(*
SPDX-FileCopyrightText: © 2026 Oleksandr Tiutyk <trofimich@gmail.com>
SPDX-License-Identifier: MIT
License: https://opensource.org/license/mit
*)

(*!
<summary>Provides static helper methods for throwing Workflow-specific exceptions.</summary>
<description>
Constructs stack-local template exceptions, formats diagnostics without heap allocation and propagates them
through ExceptionManager. Formatting uses bounded storage; propagation may allocate a registered clone.
Call only from cyclic execution, outside lifecycle methods. Each template is call-local; exception ownership
and task-boundary cleanup remain governed by Core.ExceptionManager and DynamicMemoryManager.
</description>
*)

{attribute 'no_explicit_call' := 'do not call this function block directly'}
PROGRAM WorkflowExceptions
VAR
	{attribute 'hide'} 
	_ClassName : STRING := __POUNAME();
END_VAR

(*!
<summary>Returns the diagnostic name stored by this program.</summary>
<description>
Borrows program-owned storage. Treat the returned reference as read-only and do not use it to change metadata.
</description>
*)
{attribute 'monitoring' := 'call'}
PROPERTY ClassName : REFERENCE TO STRING
GET
ClassName REF= _ClassName;
END_GET
END_PROPERTY

(*!
<summary>Returns the compiler-initialized library namespace.</summary>
<description>
Borrows shared read-only namespace storage; no allocation or ownership transfer occurs.
</description>
*)
{attribute 'monitoring' := 'call'}
PROPERTY NamespaceName : REFERENCE TO STRING
GET
NamespaceName REF= CurrentNamespace.Name;
END_GET
END_PROPERTY

(*!
<summary>Raises an InvalidNestedWorkflowStateException without requiring a caller-owned exception variable.</summary>
<description>
Constructs a temporary stack template and delegates to InvalidNestedWorkflowStateException.Throw.
</description>
<param name="sourceNamespaceName">Namespace of the caller.</param>
<param name="sourceClassName">Class name of the caller.</param>
<param name="sourcePOUName">POU name of the caller.</param>
<param name="sourcePosition">Source position of the caller.</param>
<param name="nestedActivityState">Observed child workflow element state.</param>
*)
METHOD ThrowInvalidNestedWorkflowState
VAR_INPUT
	sourceNamespaceName : STRING;
	sourceClassName : STRING;
	sourcePOUName : STRING;
	sourcePosition : STRING;
	nestedActivityState : WORKFLOW_ELEMENT_STATE;
END_VAR
VAR
	exception : InvalidNestedWorkflowStateException;
END_VAR
exception.Throw(
	sourceNamespaceName := sourceNamespaceName,
	sourceClassName := sourceClassName,
	sourcePOUName := sourcePOUName,
	sourcePosition := sourcePosition,
	nestedActivityState := nestedActivityState
);
END_METHOD

(*!
<summary>Raises an InvalidWorkflowTransitionException without requiring a caller-owned exception variable.</summary>
<description>
Constructs a temporary stack template and delegates to InvalidWorkflowTransitionException.Throw.
</description>
<param name="sourceNamespaceName">Namespace of the caller.</param>
<param name="sourceClassName">Class name of the caller.</param>
<param name="sourcePOUName">POU name of the caller.</param>
<param name="sourcePosition">Source position of the caller.</param>
<param name="fromState">Current state of the workflow element.</param>
<param name="toState">Rejected target state.</param>
*)
METHOD ThrowInvalidWorkflowTransition
VAR_INPUT
	sourceNamespaceName : STRING;
	sourceClassName : STRING;
	sourcePOUName : STRING;
	sourcePosition : STRING;
	fromState : WORKFLOW_ELEMENT_STATE;
	toState : WORKFLOW_ELEMENT_STATE;
END_VAR
VAR
	exception : InvalidWorkflowTransitionException;
END_VAR
exception.Throw(
	sourceNamespaceName := sourceNamespaceName,
	sourceClassName := sourceClassName,
	sourcePOUName := sourcePOUName,
	sourcePosition := sourcePosition,
	fromState := fromState,
	toState := toState
);
END_METHOD

(*!
<summary>Raises a WorkflowAttachmentException without requiring a caller-owned exception variable.</summary>
<description>Constructs a temporary stack template and delegates to WorkflowAttachmentException.Throw.</description>
<param name="sourceNamespaceName">Namespace of the caller.</param>
<param name="sourceClassName">Class name of the caller.</param>
<param name="sourcePOUName">POU name of the caller.</param>
<param name="sourcePosition">Source position of the caller.</param>
<param name="message">Diagnostic explanation.</param>
*)
METHOD ThrowWorkflowAttachment
VAR_INPUT
	sourceNamespaceName : STRING;
	sourceClassName : STRING;
	sourcePOUName : STRING;
	sourcePosition : STRING;
END_VAR
VAR_IN_OUT CONSTANT
	message : TOF_Core.ERROR_MESSAGE;
END_VAR
VAR
	exception : WorkflowAttachmentException;
END_VAR
exception.Throw(
	sourceNamespaceName := sourceNamespaceName,
	sourceClassName := sourceClassName,
	sourcePOUName := sourcePOUName,
	sourcePosition := sourcePosition,
	message := message
);
END_METHOD

(*!
<summary>Raises a WorkflowConfigurationException without requiring a caller-owned exception variable.</summary>
<description>Constructs a temporary stack template and delegates to WorkflowConfigurationException.Throw.</description>
<param name="sourceNamespaceName">Namespace of the caller.</param>
<param name="sourceClassName">Class name of the caller.</param>
<param name="sourcePOUName">POU name of the caller.</param>
<param name="sourcePosition">Source position of the caller.</param>
<param name="message">Diagnostic explanation.</param>
*)
METHOD ThrowWorkflowConfiguration
VAR_INPUT
	sourceNamespaceName : STRING;
	sourceClassName : STRING;
	sourcePOUName : STRING;
	sourcePosition : STRING;
	message : WSTRING(255);
END_VAR
VAR
	exception : WorkflowConfigurationException;
END_VAR
exception.Throw(
	sourceNamespaceName := sourceNamespaceName,
	sourceClassName := sourceClassName,
	sourcePOUName := sourcePOUName,
	sourcePosition := sourcePosition,
	message := message
);
END_METHOD

(*!
<summary>Raises a WorkflowVariableNotFoundException without requiring a caller-owned exception variable.</summary>
<description>
Constructs a temporary stack template and delegates to WorkflowVariableNotFoundException.Throw.
</description>
<param name="sourceNamespaceName">Namespace of the caller.</param>
<param name="sourceClassName">Class name of the caller.</param>
<param name="sourcePOUName">POU name of the caller.</param>
<param name="sourcePosition">Source position of the caller.</param>
<param name="message">Diagnostic explanation.</param>
*)
METHOD ThrowWorkflowVariableNotFound
VAR_INPUT
	sourceNamespaceName : STRING;
	sourceClassName : STRING;
	sourcePOUName : STRING;
	sourcePosition : STRING;
END_VAR
VAR_IN_OUT CONSTANT
	message : TOF_Core.ERROR_MESSAGE;
END_VAR
VAR
	exception : WorkflowVariableNotFoundException;
END_VAR
exception.Throw(
	sourceNamespaceName := sourceNamespaceName,
	sourceClassName := sourceClassName,
	sourcePOUName := sourcePOUName,
	sourcePosition := sourcePosition,
	message := message
);
END_METHOD

END_PROGRAM

(* stored: Version 1.1.0.1
   POU WorkflowExceptions: Id {66dc72bd-64d8-44a5-91d6-25d539c474f9}, SpecialFunc None
   Property ClassName: Id {794c93b6-fce0-4f75-9f7c-6316342f9fad}
   Get Get: Id {efc5ea2e-5a89-4198-aacb-5f6eb07151b0}
   Property NamespaceName: Id {639a2c56-6e40-4746-aa3c-483445eb911c}
   Get Get: Id {64a8399f-a360-4fce-ac79-db6fc38b2520}
   Method ThrowInvalidNestedWorkflowState: Id {dac3b225-92f2-4a39-b79e-295c66611eb1}
   Method ThrowInvalidWorkflowTransition: Id {07c7d49c-38ae-4a44-8d11-c642759b13f3}
   Method ThrowWorkflowAttachment: Id {2f87586b-d5f8-4b04-8ced-bda03a83e725}
   Method ThrowWorkflowConfiguration: Id {a4f608c3-b8cb-48fe-aab5-91a8b16211ab}
   Method ThrowWorkflowVariableNotFound: Id {b28ba92d-2541-49f3-a377-42842d826a53} *)
